// TIA Portal V20 export
TYPE "Störmeldung"
   STRUCT
      Störmeldung : Array[0..31] of Bool;
   END_STRUCT;
END_TYPE
